FUNCTION F_ControlDecision : UINT
// 纯仲裁判定，方便针对真实 ST 条件进行离线边界测试。
VAR_INPUT
    nOwner : UINT; // 当前控制权持有站；0 未分配，1 控制室、2 拖车本地、3 远程室。
    nStation : UINT; // 本次申请或释放的来源站号，合法范围 1～3，站号越小优先级越高。
    nAction : UINT; // 本次控制权操作：1 申请，2 释放。
    xLocked : BOOL; // 统一交接锁；TRUE 时拒绝转交或释放，持有站重复申请仍可确认授权。
    xOnline : BOOL; // 请求来源站心跳在线标志；FALSE 时拒绝该站请求。
END_VAR

// 成功应答不总表示交接：本持有者重复申请只是确认已有权限。
IF (nStation < 1) OR (nStation > 3) OR ((nAction <> 1) AND (nAction <> 2)) THEN
    F_ControlDecision := 7;
ELSIF NOT xOnline THEN
    F_ControlDecision := 4;
ELSIF (nAction = 1) AND (nOwner = nStation) THEN
    F_ControlDecision := 1;
ELSIF xLocked THEN
    // 用户规则：运行中包括高优先级站在内，不能申请接管，也不能主动释放。
    F_ControlDecision := 2;
ELSIF nAction = 2 THEN
    IF nOwner = nStation THEN F_ControlDecision := 1;
    ELSE F_ControlDecision := 5;
    END_IF
ELSIF (nOwner <> 0) AND (nStation > nOwner) THEN
    F_ControlDecision := 6;
ELSE
    F_ControlDecision := 1;
END_IF

END_FUNCTION

(* stored: Version 1.1.0.1
   POU F_ControlDecision: Id {21D9CA08-245A-44FC-B2E8-A91FE26405D0}, SpecialFunc None *)
